(* IEC 61131-3 sources: bevling_machine/framework/sources/02_Devices, 14 files *)

(* ---- F_At.st ---- *)
(* 模块说明：检查设备可用、无忙无故障且位置误差小于 0.01。它检查位置，不检查本次命令序号。 *)
FUNCTION F_At : BOOL
VAR_INPUT
    stStatus : ST_DeviceStatus; (* 本模块对外发布的状态；字段含义见其数据类型。 *)
    lrTarget : LREAL; (* 要检查的目标位置；误差小于 0.01 且设备就绪、无忙无错时返回 TRUE。 *)
END_VAR
FUNCTION F_At : BOOL
(* 位置容差为 0.01 工程单位；这里不做新命令序号校验，用于姿态/互锁判断。 *)
F_At := stStatus.xReady AND NOT stStatus.xBusy
    AND NOT stStatus.xError AND (ABS(stStatus.lrPosition-lrTarget) < 0.01);

(* ---- F_Command.st ---- *)
(* 模块说明：组装设备命令，不执行运动。由设备管理器和对应设备功能块实际处理。 *)
FUNCTION F_Command : ST_DeviceCommand
VAR_INPUT
    eAction : E_DeviceAction; (* 动作类型：无请求、定位、连续运行、点动或停止，见 E_DeviceAction。 *)
    udiID : UDINT; (* 本次命令序号，0 无效；发起新定位时换新序号。 *)
    lrTarget : LREAL; (* 目标工程位置；气缸使用约定的 0/1 端点，连续运行和点动不使用该位置。 *)
    lrVelocity : LREAL; (* 请求速度，单位随设备工程单位定义；尚未完成实机标定。 *)
END_VAR
FUNCTION F_Command : ST_DeviceCommand
(* 只复制字段形成结构体，不等待动作、不直接访问物理设备。 *)
F_Command.eAction := eAction;
F_Command.udiID := udiID;
F_Command.lrTarget := lrTarget;
F_Command.lrVelocity := lrVelocity;

(* ---- F_Done.st ---- *)
(* 模块说明：只有设备完成序号等于本次命令序号、无忙且无故障，才返回动作完成。 *)
FUNCTION F_Done : BOOL
VAR_INPUT
    stStatus : ST_DeviceStatus; (* 本模块对外发布的状态；字段含义见其数据类型。 *)
    udiID : UDINT; (* 本次命令序号，0 无效；发起新定位时换新序号。 *)
END_VAR
FUNCTION F_Done : BOOL
(* 完成必须匹配本次请求；历史 Done 或仅 Busy=FALSE 都不足以作为本步完成条件。 *)
F_Done := (udiID <> 0) AND (stStatus.udiCompletedID = udiID)
    AND NOT stStatus.xBusy AND NOT stStatus.xError;

(* ---- F_NextID.st ---- *)
(* 模块说明：生成本次动作的非零序号。计数到最大值后回到 1，用于排除上一步残留的完成反馈。 *)
FUNCTION F_NextID : UDINT
VAR_IN_OUT
    udiCounter : UDINT; (* 全机共享的动作序号计数器，通过引用传递；由 F_NextID 分配，0 不使用。 *)
END_VAR
FUNCTION F_NextID : UDINT
(* 最大值之后回到 1，跳过无效序号 0；同一机台所有流程共享该计数器。 *)
IF udiCounter = 16#FFFFFFFF THEN udiCounter := 1;
ELSE udiCounter := udiCounter + 1;
END_IF
F_NextID := udiCounter;

(* ---- F_SafetyBypassActive.st ---- *)
(* 模块说明：安全许可软件旁路的唯一判定点。两级开关同时置位才返回 TRUE。 *)
FUNCTION F_SafetyBypassActive : BOOL
VAR_IN_OUT
	stReal : ST_RealDeviceSettings; (* 引用传递，避免每次扫描拷贝整个设置结构体。 *)
END_VAR
FUNCTION F_SafetyBypassActive : BOOL
(* 一级开关与二级确认必须同时置位；任一为 FALSE 就返回 FALSE，保持原有安全逻辑。 *)
F_SafetyBypassActive := stReal.xSafetyBypass AND stReal.xSafetyBypassConfirm;

(* ---- FB_Axis.st ---- *)
(* 模块说明：定位轴适配入口。当前调用内部仿真；真实轴的 MC 功能块、回原点和限位尚未接入。 *)
FUNCTION_BLOCK FB_Axis
VAR_INPUT
    xSimulation : BOOL; (* TRUE 使用内部仿真；当前 FALSE 报未实现 3001，不会接管真实运动。 *)
    xEnable : BOOL; (* 本功能使能，电平有效；失能时不接受新的动作请求。 *)
    xReset : BOOL; (* 故障复位许可；仿真设备仅在故障注入已撤销时清除错误。 *)
    xStall : BOOL; (* 仿真卡住输入；TRUE 暂停位置推进且不发完成，保留忙状态。 *)
    xInjectFault : BOOL; (* 仿真设备故障输入；TRUE 锁存错误码 9001。 *)
    stConfig : ST_DeviceConfig; (* 设备类型、初始位置、软限位与仿真动作时间。 *)
    stCommand : ST_DeviceCommand; (* 当前单设备命令，含动作类型、序号、目标和速度。 *)
END_VAR
VAR_OUTPUT
    stStatus : ST_DeviceStatus; (* 本模块对外发布的状态；字段含义见其数据类型。 *)
END_VAR
VAR
    fbSimulation : FB_SimDevice; (* 内部设备仿真实例，真实设备适配尚未接入。 *)
END_VAR
FUNCTION_BLOCK FB_Axis
(* 真实设备适配尚未接入；关闭仿真时返回 3001，避免误认为已具备实机控制。 *)
fbSimulation(xEnable := xEnable AND xSimulation, xReset := xReset,
    xStall := xStall, xInjectFault := xInjectFault,
    stConfig := stConfig, stCommand := stCommand);
stStatus := fbSimulation.stStatus;
IF NOT xSimulation THEN
    stStatus.xReady := FALSE; stStatus.xBusy := FALSE; stStatus.xActive := FALSE;
    stStatus.xError := TRUE; stStatus.udiErrorID := 3001;
END_IF

(* ---- FB_Cylinder.st ---- *)
(* 模块说明：气缸适配入口。当前用 0/1 位置模拟两端到位；真实电磁阀和到位传感器尚未映射。 *)
FUNCTION_BLOCK FB_Cylinder
VAR_INPUT
    xSimulation : BOOL; (* TRUE 使用内部仿真；当前 FALSE 报未实现 3001，不会接管真实运动。 *)
    xEnable : BOOL; (* 本功能使能，电平有效；失能时不接受新的动作请求。 *)
    xReset : BOOL; (* 故障复位许可；仿真设备仅在故障注入已撤销时清除错误。 *)
    xStall : BOOL; (* 仿真卡住输入；TRUE 暂停位置推进且不发完成，保留忙状态。 *)
    xInjectFault : BOOL; (* 仿真设备故障输入；TRUE 锁存错误码 9001。 *)
    stConfig : ST_DeviceConfig; (* 设备类型、初始位置、软限位与仿真动作时间。 *)
    stCommand : ST_DeviceCommand; (* 当前单设备命令，含动作类型、序号、目标和速度。 *)
END_VAR
VAR_OUTPUT
    stStatus : ST_DeviceStatus; (* 本模块对外发布的状态；字段含义见其数据类型。 *)
END_VAR
VAR
    fbSimulation : FB_SimDevice; (* 内部设备仿真实例，真实设备适配尚未接入。 *)
END_VAR
FUNCTION_BLOCK FB_Cylinder
(* 真实设备适配尚未接入；关闭仿真时返回 3001，避免误认为已具备实机控制。 *)
fbSimulation(xEnable := xEnable AND xSimulation, xReset := xReset,
    xStall := xStall, xInjectFault := xInjectFault,
    stConfig := stConfig, stCommand := stCommand);
stStatus := fbSimulation.stStatus;
IF NOT xSimulation THEN
    stStatus.xReady := FALSE; stStatus.xBusy := FALSE; stStatus.xActive := FALSE;
    stStatus.xError := TRUE; stStatus.udiErrorID := 3001;
END_IF

(* ---- FB_DeviceManager.st ---- *)
FUNCTION_BLOCK FB_DeviceManager
(* 模块说明：统一设备执行入口。首次建立类型和初始位置，每扫描周期按类型调用设备功能块并收集反馈。 *)
VAR_INPUT
	xEnable : BOOL; (* 本功能使能，电平有效；失能时不接受新的动作请求。 *)
	xSimulation : BOOL; (* TRUE 使用内部仿真；当前 FALSE 报未实现 3001，不会接管真实运动。 *)
	xReset : BOOL; (* 故障复位许可；仿真设备仅在故障注入已撤销时清除错误。 *)
	xFaultHold : BOOL; (* 整机故障保持：TRUE 时真实轴强制停车、真实阀失电，直到复位。 *)
	stSim : ST_SimulationSettings; (* 软件仿真设置；设备管理器按设备索引读取卡住与故障注入。 *)
	stReal : ST_RealDeviceSettings; (* 真实设备接管设置；逐台位决定该编号走真实轴还是仿真。 *)
	uiMaterialModel : UINT; (* 当前运行料型 300/450/600；G2 气缸组按此选通其中一个缸下降。 *)
	aCommand : ARRAY[1..17] OF ST_DeviceCommand; (* 统一设备请求数组 1..17；子流程写请求，设备管理器执行。 *)
END_VAR
VAR_OUTPUT
	aStatus : ARRAY[1..17] OF ST_DeviceStatus; (* 各设备的反馈数组 1..17，供判断忙、完成序号、故障和位置。 *)
	aValveOut : ARRAY[1..17] OF BOOL; (* 各设备的阀电气输出电平 1..17；只有已接管的真实气缸可能为 TRUE，供物理映射层取用。 *)
	aValveOutAux : ARRAY[1..17] OF BOOL; (* 第二个执行器的阀电气电平 1..17；当前只有 G1 双压板的 [9] 有效，其余恒 FALSE。 *)
	aG2Valve : ARRAY[1..3] OF BOOL; (* G2 三个侧挡阀的电气电平 1=300，2=450，3=600；未接管时全 FALSE。 *)
	uiG2Band : UINT; (* G2 当前实际下降的料型带号 300/450/600；0 表示三缸全部提升，供诊断观察。 *)
END_VAR
VAR
	aConfig : ARRAY[1..17] OF ST_DeviceConfig; (* 设备配置数组，首扫描按固定编号设置类型和初始姿态。 *)
	aAxis : ARRAY[1..17] OF FB_Axis; (* 定位轴功能块实例数组，只有设备类型为 Axis 的元素被调用。 *)
	aMotor : ARRAY[1..17] OF FB_Motor; (* 连续电机功能块实例数组，供 D1、D3 使用。 *)
	aCylinder : ARRAY[1..17] OF FB_Cylinder; (* 气缸功能块实例数组，按 G 编号驱动对应仿真实例。 *)
	aValve : ARRAY[1..17] OF FB_Valve; (* 阀功能块实例数组，供 G5 喷油及 G6 吹气使用。 *)
	fbRealD1 : FB_RealAxis; (* D1 送料皮带真实轴实例，绑定 songliao。 *)
	fbRealD2 : FB_RealAxis; (* D2 切割走刀真实轴实例，绑定 qiege。 *)
	fbRealD3 : FB_RealAxis; (* D3 盘刀旋转真实轴实例，绑定 pandao（当前按线性模式配置）。 *)
	fbRealD8 : FB_RealAxis; (* D8 平台旋转真实轴实例，绑定 xuanzhuan（台达 ASDA-B3-E）。 *)
	fbRealG1 : FB_RealCylinder; (* G1 下压气缸真实实例，绑定左右两路阀与 G1 两端传感器。 *)
	fbRealG2 : FB_RealCylinderGroup; (* G2 侧挡气缸组真实实例，一台管 300/450/600 三个缸。 *)
	fbRealG3 : FB_RealCylinder; (* G3 侧推气缸真实实例，绑定 xDoG3Valve 与 G3 两端传感器。 *)
	fbRealG9 : FB_RealCylinder; (* G9 盘刀升降真实实例，绑定 xDoG9Valve 与 G9 两端传感器。 *)
	fbRealD6 : FB_RealSensor; (* D6 定长光电真实实例，只读；接管后取代 FB_SimPlant 产生料到位信号。 *)
	axUseReal : ARRAY[1..17] OF BOOL; (* 本扫描逐台接管标志，直接取 stReal.axRealDevice；没有真实实例的编号由回填分支报 3002。 *)
	xBooted : BOOL; (* 本功能块首次初始化完成标志，防止每扫描重写初值。 *)
	i : INT; (* 本扫描数组遍历索引；含义及范围以当前 FOR 循环为准。 *)
END_VAR
FUNCTION_BLOCK FB_DeviceManager
IF NOT xBooted THEN
	(* D1 送料皮带：由真实轴 songliao 承担输送，按定位轴建模（点动/连续运行）。 *)
	aConfig[1].eKind := E_DeviceKind.Axis;
	aConfig[2].eKind := E_DeviceKind.Axis;
	aConfig[3].eKind := E_DeviceKind.Motor;
	aConfig[4].eKind := E_DeviceKind.Axis;
	(* D5 暂按定位升降建模：0=升起避让，1=下降检测，非实际机械坐标。 *)
	aConfig[5].eKind := E_DeviceKind.Axis;
	aConfig[7].eKind := E_DeviceKind.Axis;
	aConfig[8].eKind := E_DeviceKind.Axis;
	FOR i := 9 TO 17 DO aConfig[i].eKind := E_DeviceKind.Cylinder; END_FOR
	aConfig[13].eKind := E_DeviceKind.Valve;
	aConfig[14].eKind := E_DeviceKind.Valve;
	aConfig[12].lrInitialPosition := 1.0;
	FOR i := 1 TO 17 DO
		IF aConfig[i].eKind = E_DeviceKind.Cylinder THEN
			aConfig[i].lrMinPosition := 0.0; aConfig[i].lrMaxPosition := 1.0;
		END_IF
	END_FOR
	(* D2 切割走刀：配方要求 200mm/s、加速度 500；默认 100/50 会把速度削到 100 并拖长加减速段。 *)
	aConfig[2].lrMaxVelocity := 300.0;
	aConfig[2].lrMaxAcceleration := 500.0;
	aConfig[2].lrMaxDeceleration := 500.0;
	xBooted := TRUE;
END_IF

(* 逐台接管标志直接取设置位：是否真的接管由下方回填分支的 CASE 决定。
   新增真实实例时只改 CASE 和实例调用两处，不要再维护第二份白名单。 *)
FOR i := 1 TO 17 DO
	axUseReal[i] := stReal.axRealDevice[i];
END_FOR

(* 四个真实轴实例每扫描必须无条件调用；轴形参写死，无法放进 FOR 循环。
   绑定对照（换电机、改轴名后必须逐行核对：写错不会报编译错误，
   因为任何一个合法轴名都能通过类型检查，只能靠单点测试发现）：
     fbRealD1 -> songliao    设备索引 1，送料皮带（EtherCAT 从站 ASDA_B3_E_CoE_Drive_3）
     fbRealD2 -> qiege       设备索引 2，切割走刀（从站 ASDA_B3_E_CoE_Drive_1）
     fbRealD3 -> pandao      设备索引 3，盘刀旋转（从站 ASDA_B3_E_CoE_Drive_2）
     fbRealD8 -> xuanzhuan   设备索引 8，平台旋转（从站 ASDA_B3_E_CoE_Drive，台达）
   注意：ASDA_B3_E_CoE_Drive_* 是驱动器从站名，代码里写的必须是它下面那个
   轴对象名（songliao/qiege/pandao/xuanzhuan），两者不是一回事。 *)
fbRealD1(Axis := songliao, xUseReal := axUseReal[1], xEnable := xEnable, xReset := xReset,
	xFaultHold := xFaultHold,
	stConfig := aConfig[1], stCommand := aCommand[1], stReal := stReal);
fbRealD2(Axis := qiege, xUseReal := axUseReal[2], xEnable := xEnable, xReset := xReset,
	xFaultHold := xFaultHold,
	stConfig := aConfig[2], stCommand := aCommand[2], stReal := stReal);
fbRealD3(Axis := pandao, xUseReal := axUseReal[3], xEnable := xEnable, xReset := xReset,
	xFaultHold := xFaultHold,
	stConfig := aConfig[3], stCommand := aCommand[3], stReal := stReal);
fbRealD8(Axis := xuanzhuan, xUseReal := axUseReal[8], xEnable := xEnable, xReset := xReset,
	xFaultHold := xFaultHold,
	stConfig := aConfig[8], stCommand := aCommand[8], stReal := stReal);

(* 四个真实气缸实例同样必须无条件调用；传感器与阀逐一对应物理映射符号。
   极性默认 FALSE：传感器高电平有效、阀高电平使能。接线反了只改这里一行，不动流程与互锁。 *)
fbRealG1(xUseReal := axUseReal[9], xEnable := xEnable, xReset := xReset,
	xFaultHold := xFaultHold,
	xSensorRetract := GVL_IO_Physical.xDiG1LRetract, xSensorExtend := GVL_IO_Physical.xDiG1LExtend,
	xSensorRetract2 := GVL_IO_Physical.xDiG1RRetract, xSensorExtend2 := GVL_IO_Physical.xDiG1RExtend,
	xUseSecond := TRUE,
	(* 现场 G1 两只伸出到位传感器已失效：改成只看左右两个缩回信号，两者都无信号并稳定 1s 即认为压到位。
	   传感器修好后把 xExtendByRetract 改回 FALSE 就恢复两端判定，流程和互锁都不用动。 *)
	xExtendByRetract := TRUE, tExtendConfirm := T#1S,
	xInvertSensors := FALSE, xInvertValve := FALSE,
	stConfig := aConfig[9], stCommand := aCommand[9]);
fbRealG2(xUseReal := axUseReal[10], xEnable := xEnable, xReset := xReset,
	xFaultHold := xFaultHold,
	uiMaterialModel := uiMaterialModel,
	xSensorRetract1 := GVL_IO_Physical.xDiG2_300Retract, xSensorExtend1 := GVL_IO_Physical.xDiG2_300Extend,
	xSensorRetract2 := GVL_IO_Physical.xDiG2_450Retract, xSensorExtend2 := GVL_IO_Physical.xDiG2_450Extend,
	xSensorRetract3 := GVL_IO_Physical.xDiG2_600Retract, xSensorExtend3 := GVL_IO_Physical.xDiG2_600Extend,
	xInvertSensors := FALSE, xInvertValve := FALSE,
	stConfig := aConfig[10], stCommand := aCommand[10]);
fbRealG3(xUseReal := axUseReal[11], xEnable := xEnable, xReset := xReset,
	xFaultHold := xFaultHold,
	xSensorRetract := GVL_IO_Physical.xDiG3Retract, xSensorExtend := GVL_IO_Physical.xDiG3Extend,
	xInvertSensors := FALSE, xInvertValve := FALSE,
	stConfig := aConfig[11], stCommand := aCommand[11]);
fbRealG9(xUseReal := axUseReal[17], xEnable := xEnable, xReset := xReset,
	xFaultHold := xFaultHold,
	xSensorRetract := GVL_IO_Physical.xDiG9Retract, xSensorExtend := GVL_IO_Physical.xDiG9Extend,
	xInvertSensors := FALSE, xInvertValve := FALSE,
	stConfig := aConfig[17], stCommand := aCommand[17]);

(* D6 定长光电：只读设备，没有阀也没有动作。
   接线极性反了改 xInvertSensor；光电抖动大改 tDebounce；不需要常亮/常灭监视就把 tStuckTimeout 置 T#0MS。 *)
fbRealD6(xUseReal := axUseReal[6], xEnable := xEnable, xReset := xReset,
	xSensorRaw := GVL_IO_Physical.xDiMaterialLength, xInvertSensor := FALSE,
	tDebounce := T#20MS, tStuckTimeout := T#0MS,
	stConfig := aConfig[6], stCommand := aCommand[6]);

(* 每周期按接管标志二选一：有真实实例的直接回填，否则按设备类型走仿真。
   「实例即事实」：本 CASE 列出全部已实现真实适配的编号，没列到的编号若置了接管位，
   就在 ELSE 分支明确报 3002，避免静默走仿真被误认为已接实机。 *)
(* G2 三个阀默认失电：只有走真实气缸组且缸确实在下降时才会被下面的 CASE 置位。 *)
aG2Valve[1] := FALSE; aG2Valve[2] := FALSE; aG2Valve[3] := FALSE;
uiG2Band := 0;
FOR i := 1 TO 17 DO
	aValveOut[i] := FALSE; aValveOutAux[i] := FALSE;
	IF axUseReal[i] THEN
		CASE i OF
		1: aStatus[i] := fbRealD1.stStatus;
		2: aStatus[i] := fbRealD2.stStatus;
		3: aStatus[i] := fbRealD3.stStatus;
		6: aStatus[i] := fbRealD6.stStatus;
		8: aStatus[i] := fbRealD8.stStatus;
		9: aStatus[i] := fbRealG1.stStatus; aValveOut[i] := fbRealG1.xValve; aValveOutAux[i] := fbRealG1.xValve2;
		10: aStatus[i] := fbRealG2.stStatus; aG2Valve := fbRealG2.aValve; uiG2Band := fbRealG2.uiActiveBand;
		11: aStatus[i] := fbRealG3.stStatus; aValveOut[i] := fbRealG3.xValve;
		17: aStatus[i] := fbRealG9.stStatus; aValveOut[i] := fbRealG9.xValve;
		ELSE
			(* 请求接管但本版本没有对应真实实例：只报错，不启动仿真，保持与老逻辑一致 *)
			aStatus[i].xError := TRUE;
			aStatus[i].udiErrorID := 3002;
		END_CASE
	ELSE
		CASE aConfig[i].eKind OF
		E_DeviceKind.Axis:
			aAxis[i](xSimulation:=xSimulation,xEnable:=xEnable,xReset:=xReset,
				xStall:=stSim.axStall[i],xInjectFault:=stSim.axFault[i],stConfig:=aConfig[i],stCommand:=aCommand[i]);
			aStatus[i] := aAxis[i].stStatus;
		E_DeviceKind.Motor:
			aMotor[i](xSimulation:=xSimulation,xEnable:=xEnable,xReset:=xReset,
				xStall:=stSim.axStall[i],xInjectFault:=stSim.axFault[i],stConfig:=aConfig[i],stCommand:=aCommand[i]);
			aStatus[i] := aMotor[i].stStatus;
		E_DeviceKind.Cylinder:
			aCylinder[i](xSimulation:=xSimulation,xEnable:=xEnable,xReset:=xReset,
				xStall:=stSim.axStall[i],xInjectFault:=stSim.axFault[i],stConfig:=aConfig[i],stCommand:=aCommand[i]);
			aStatus[i] := aCylinder[i].stStatus;
		E_DeviceKind.Valve:
			aValve[i](xSimulation:=xSimulation,xEnable:=xEnable,xReset:=xReset,
				xStall:=stSim.axStall[i],xInjectFault:=stSim.axFault[i],stConfig:=aConfig[i],stCommand:=aCommand[i]);
			aStatus[i] := aValve[i].stStatus;
		END_CASE
	END_IF
END_FOR

(* ---- FB_Motor.st ---- *)
(* 模块说明：连续电机适配入口，供皮带 D1 和盘刀 D3 使用。当前仅仿真运行状态。 *)
FUNCTION_BLOCK FB_Motor
VAR_INPUT
    xSimulation : BOOL; (* TRUE 使用内部仿真；当前 FALSE 报未实现 3001，不会接管真实运动。 *)
    xEnable : BOOL; (* 本功能使能，电平有效；失能时不接受新的动作请求。 *)
    xReset : BOOL; (* 故障复位许可；仿真设备仅在故障注入已撤销时清除错误。 *)
    xStall : BOOL; (* 仿真卡住输入；TRUE 暂停位置推进且不发完成，保留忙状态。 *)
    xInjectFault : BOOL; (* 仿真设备故障输入；TRUE 锁存错误码 9001。 *)
    stConfig : ST_DeviceConfig; (* 设备类型、初始位置、软限位与仿真动作时间。 *)
    stCommand : ST_DeviceCommand; (* 当前单设备命令，含动作类型、序号、目标和速度。 *)
END_VAR
VAR_OUTPUT
    stStatus : ST_DeviceStatus; (* 本模块对外发布的状态；字段含义见其数据类型。 *)
END_VAR
VAR
    fbSimulation : FB_SimDevice; (* 内部设备仿真实例，真实设备适配尚未接入。 *)
END_VAR
FUNCTION_BLOCK FB_Motor
(* 真实设备适配尚未接入；关闭仿真时返回 3001，避免误认为已具备实机控制。 *)
fbSimulation(xEnable := xEnable AND xSimulation, xReset := xReset,
    xStall := xStall, xInjectFault := xInjectFault,
    stConfig := stConfig, stCommand := stCommand);
stStatus := fbSimulation.stStatus;
IF NOT xSimulation THEN
    stStatus.xReady := FALSE; stStatus.xBusy := FALSE; stStatus.xActive := FALSE;
    stStatus.xError := TRUE; stStatus.udiErrorID := 3001;
END_IF

(* ---- FB_RealAxis.st ---- *)
FUNCTION_BLOCK FB_RealAxis
(* 模块说明：真实轴适配层。把统一设备命令翻译成 SoftMotion 动作，并回写与仿真完全一致的接收/完成序号。 *)
VAR_IN_OUT
	Axis : AXIS_REF_SM3; (* 轴节点引用，编译期强制绑定；未接轴无法通过编译，不存在空指针。 *)
END_VAR
VAR_INPUT
	xUseReal : BOOL; (* TRUE 表示本编号由本功能块接管；FALSE 时驱动器保持去使能且不响应任何命令。 *)
	xEnable : BOOL; (* 设备级使能，来自整机许可；FALSE 时主动停止并清序号。 *)
	xReset : BOOL; (* 故障复位，上升沿清锁存错误与 MC 错误。 *)
	stConfig : ST_DeviceConfig; (* 行程、速度、加减速与绝对定位许可。 *)
	stCommand : ST_DeviceCommand; (* 上层统一设备命令，含义与仿真侧完全一致。 *)
	xFaultHold : BOOL; (* 整机故障保持：TRUE 期间强制 MC_Stop 常置并清所有运动请求，直到复位。 *)
	stReal : ST_RealDeviceSettings; (* 相对验证距离、速度与旁路设置。 *)
END_VAR
VAR_OUTPUT
	stStatus : ST_DeviceStatus; (* 与 FB_SimDevice 语义一致，上层无需区分真假设备。 *)
	uiVerifyPhase : UINT; (* 相对验证相位：0 空闲、1 正向、2 停留、3 反向、4 完成、90 中止。 *)
	lrVerifyMeasured : LREAL; (* 本次往返正向段的实测位移，取自轴反馈。 *)
	lrVerifyRatio : LREAL; (* 实测除以指令；只能证明指令与反馈自洽，不能证明单位就是毫米。 *)
END_VAR
VAR
	fbPower : MC_Power; (* 伺服使能，接管期间保持上电。 *)
	fbReset : MC_Reset; (* 清 MC 错误。 *)
	fbStop : MC_Stop; (* 受控停止，停止请求需保持到 Done。 *)
	fbMoveAbs : MC_MoveAbsolute; (* 绝对定位，仅在 xAbsoluteAllowed 为 TRUE 时使用。 *)
	fbMoveRel : MC_MoveRelative; (* 相对定位，验证模式的两段行程使用。 *)
	fbMoveVel : MC_MoveVelocity; (* 连续运行与点动共用，两者相位互斥；方向必须显式给出。 *)
	fbHoming : CmpHCMotion.MC_Homing; (* 上位机回零：由 PLC 自己按轴配置的回零方式走，不依赖驱动器支持 DS402 回零。 *)
	fbReadPos : MC_ReadActualPosition; (* 实际位置反馈。 *)
	fbReadStatus : MC_ReadStatus; (* 轴状态，用于判断故障停止。 *)
	fbReadErr : MC_ReadAxisError; (* 轴错误码，供在线排查。 *)
	rtReset : R_TRIG; (* 复位上升沿。 *)
	tonEnable : TON; (* 命令已接收但轴未使能的 3 秒超时。 *)
	tonDwell : TON; (* 验证往返之间的停留，保证 Execute 拉低形成新上升沿。 *)
	tonHome : TON; (* 回零超时；找不到原点时按 2004 暴露，避免无限等待。 *)
	udiLastID : UDINT; (* 上次已接受序号，用于识别新命令。 *)
	udiActiveID : UDINT; (* 正在执行的序号，完成时回写。 *)
	xPending : BOOL; (* 已接收但尚未启动，等待轴使能。 *)
	xStopLatch : BOOL; (* 停止请求锁存，保持到 MC_Stop 完成。 *)
	xStopReq : BOOL; (* 本扫描停止请求。 *)
	xMoveAbsReq : BOOL; (* 本扫描绝对定位请求。 *)
	xMoveRelReq : BOOL; (* 本扫描相对定位请求。 *)
	xMoveVelReq : BOOL; (* 本扫描速度模式请求，连续运行与点动共用。 *)
	xHomeReq : BOOL; (* 本扫描回零请求，保持到 Done。 *)
	xHomed : BOOL; (* 本次上电后已成功回零；成功后允许绝对定位，断电或重新下载后清零。 *)
	uiPhase : UINT; (* 动作相位：0 空闲、10 等待使能、20 绝对、30/31/32 验证三段、40 连续、50 点动、60 回零、90 中止。 *)
	lrVerifyStart : LREAL; (* 验证正向段起点位置。 *)
	lrRelDistance : LREAL; (* 本次相对定位距离，正负决定方向。 *)
	lrRelVelocity : LREAL; (* 本次相对定位速度，取正值。 *)
	lrCmdVelocity : LREAL; (* 连续运行与点动的限幅后速度，带符号。 *)
END_VAR
FUNCTION_BLOCK FB_RealAxis
(* ===== 1. 读取块无条件调用，保证反馈新鲜 ===== *)
fbReadPos(Axis := Axis, Enable := TRUE);
fbReadStatus(Axis := Axis, Enable := TRUE);
fbReadErr(Axis := Axis, Enable := TRUE);
rtReset(CLK := xReset);

stStatus.lrPosition := fbReadPos.Position;
stStatus.xRealActive := xUseReal;

(* ===== 2. 复位：只在接管状态下响应，避免误清其它轴 ===== *)
IF xUseReal AND rtReset.Q THEN
	stStatus.xError := FALSE;
	stStatus.udiErrorID := 0;
	xStopLatch := FALSE;
	xPending := FALSE;
	uiPhase := 0;
	uiVerifyPhase := 0;
	udiLastID := 0;
	udiActiveID := 0;
	stStatus.udiAcceptedID := 0;
	stStatus.udiCompletedID := 0;
	stStatus.xBusy := FALSE;
	stStatus.xActive := FALSE;
END_IF

(* ===== 3. 定时器：用上扫描状态驱动，避免与状态判定循环依赖 ===== *)
tonEnable(IN := xPending AND xUseReal, PT := T#3S);
tonDwell(IN := (uiPhase = 31), PT := stReal.tVerifyDwell);
tonHome(IN := (uiPhase = 60), PT := stReal.tHomeTimeout);

(* ===== 4. 请求默认全部撤销 ===== *)
xStopReq := FALSE;
xMoveAbsReq := FALSE;
xMoveRelReq := FALSE;
xMoveVelReq := FALSE;
xHomeReq := FALSE;
lrRelDistance := 0.0;
lrRelVelocity := 0.0;
lrCmdVelocity := 0.0;

(* ===== 4.5 整机故障保持：故障期间主动停车，不依赖 xPermit 间接撤销 ===== *)
(* 为什么需要：进入 Fault 时上层只是让 xPermit 变 FALSE，请求被换成 Stop。但 Stop 是
   一次性的动作请求，盘刀这类连续运行设备在 MC_Stop 完成后再无后续指令，表现就是
   “PLC 认为已停、实际还在转”。这里改用 xFaultHold 强制 MC_Stop 常置，直到真正复位。 *)
IF xFaultHold THEN
	xStopReq := TRUE;
	xPending := FALSE;
	xMoveAbsReq := FALSE; xMoveRelReq := FALSE; xMoveVelReq := FALSE; xHomeReq := FALSE;
	uiPhase := 0; uiVerifyPhase := 0;
	udiLastID := 0; udiActiveID := 0;
	stStatus.udiAcceptedID := 0; stStatus.udiCompletedID := 0;
	stStatus.xBusy := FALSE; stStatus.xActive := FALSE;
END_IF

(* ===== 5. 主状态判定 ===== *)
IF NOT xUseReal THEN
	(* 未接管：不产生任何运动请求，驱动器由 MC_Power 去使能。 *)
	xPending := FALSE; xStopLatch := FALSE;
	uiPhase := 0; uiVerifyPhase := 0;
	udiLastID := 0; udiActiveID := 0;
	stStatus.xReady := FALSE;
	stStatus.xBusy := FALSE; stStatus.xActive := FALSE;
	stStatus.udiAcceptedID := 0; stStatus.udiCompletedID := 0;
	stStatus.xError := FALSE; stStatus.udiErrorID := 0;
ELSIF xFaultHold THEN
	(* 故障保持：只允许停止，不接收新命令，也不发布就绪。 *)
	stStatus.xReady := FALSE;
	stStatus.xBusy := FALSE; stStatus.xActive := FALSE;
	stStatus.udiAcceptedID := 0; stStatus.udiCompletedID := 0;
ELSE
	(* --- 5.1 接收新序号：新序号就是新命令，不用边沿检测 --- *)
	IF (stCommand.udiID <> 0) AND (stCommand.udiID <> udiLastID)
		AND xEnable AND NOT stStatus.xError THEN
		udiLastID := stCommand.udiID;
		udiActiveID := udiLastID;
		stStatus.udiAcceptedID := udiActiveID;
		stStatus.udiCompletedID := 0;
		stStatus.xBusy := TRUE; stStatus.xActive := FALSE;
		uiVerifyPhase := 0;
		xPending := TRUE;
		uiPhase := 10;
		xStopLatch := FALSE;
	END_IF

	(* --- 5.2 停止请求锁存：保持到 MC_Stop 完成，不能提前撤 Execute --- *)
	IF (stCommand.eAction = E_DeviceAction.Stop) OR (NOT xEnable) THEN
		(* 只在真的有动作时才锁存，避免 Stop 常驻时每扫描重复触发 MC_Stop。 *)
		IF xPending OR (uiPhase <> 0) THEN xStopLatch := TRUE; END_IF
	ELSIF (stCommand.eAction = E_DeviceAction.None) AND (uiPhase <> 0) THEN
		xStopLatch := TRUE;
	END_IF
	IF fbStop.Done THEN xStopLatch := FALSE; END_IF

	IF xStopLatch THEN
		xStopReq := TRUE;
		xPending := FALSE;
		uiPhase := 0; uiVerifyPhase := 0;
		udiLastID := 0; udiActiveID := 0;
		stStatus.udiAcceptedID := 0; stStatus.udiCompletedID := 0;
		stStatus.xBusy := FALSE; stStatus.xActive := FALSE;
	ELSIF xPending THEN
		(* --- 5.3 等轴使能；就绪后按动作类型进入相位，3 秒未使能报 2003 --- *)
		IF fbPower.Status THEN
			xPending := FALSE;
			CASE stCommand.eAction OF
			E_DeviceAction.Position:
				(* 已回零优先走绝对定位：相对验证只是未回零时的临时替代，回零成功后不再需要。 *)
				IF xHomed OR stConfig.xAbsoluteAllowed THEN
					uiPhase := 20;
				ELSIF stReal.xRelativeVerify THEN
					lrVerifyStart := fbReadPos.Position;
					uiPhase := 30; uiVerifyPhase := 1;
				ELSE
					(* 未回零不允许绝对定位：报 2002 且不置完成位，由上层按步号超时暴露。 *)
					stStatus.xError := TRUE; stStatus.udiErrorID := 2002;
					uiPhase := 0; uiVerifyPhase := 0;
				END_IF
			E_DeviceAction.Run:
				uiPhase := 40;
			E_DeviceAction.Jog:
				uiPhase := 50;
			E_DeviceAction.Home:
				uiPhase := 60;
			ELSE
				uiPhase := 0;
			END_CASE
		ELSIF tonEnable.Q THEN
			xPending := FALSE; uiPhase := 0;
			stStatus.xError := TRUE; stStatus.udiErrorID := 2003;
			stStatus.xBusy := FALSE;
		END_IF
	END_IF

	(* --- 5.4 按相位生成限幅后的运动参数 --- *)
	CASE uiPhase OF
	30:
		lrRelDistance := LIMIT(0.0, stReal.lrVerifyDistance, 20.0);
		lrRelVelocity := LIMIT(0.01, stReal.lrVerifyVelocity, stConfig.lrMaxVelocity);
	32:
		lrRelDistance := -LIMIT(0.0, stReal.lrVerifyDistance, 20.0);
		lrRelVelocity := LIMIT(0.01, stReal.lrVerifyVelocity, stConfig.lrMaxVelocity);
	40:
		(* 连续运行：按设备配置限幅，不使用验证低速。 *)
		lrCmdVelocity := LIMIT(-stConfig.lrMaxVelocity, stCommand.lrVelocity, stConfig.lrMaxVelocity);
	50:
		(* 点动：用设备最大速度与手动上限 lrManualVelocityMax 的较小者限幅；不能再用验证速度，否则手动最高只有 2mm/s。 *)
		lrCmdVelocity := LIMIT(0.01, ABS(stCommand.lrVelocity),
			MIN(stConfig.lrMaxVelocity, stReal.lrManualVelocityMax));
		IF stCommand.lrVelocity < 0.0 THEN lrCmdVelocity := -lrCmdVelocity; END_IF
	END_CASE

	xMoveAbsReq := (uiPhase = 20);
	xMoveRelReq := (uiPhase = 30) OR (uiPhase = 32);
	xMoveVelReq := (uiPhase = 40) OR (uiPhase = 50);
	xHomeReq := (uiPhase = 60);
END_IF

(* ===== 6. MC 块无条件调用：漏调用会报 SMC_FB_WASNT_CALLED_DURING_MOTION ===== *)
fbPower(Axis := Axis, Enable := xUseReal AND xEnable,
	bRegulatorOn := xUseReal AND xEnable, bDriveStart := xUseReal AND xEnable);
fbReset(Axis := Axis, Execute := xUseReal AND rtReset.Q);
fbStop(Axis := Axis, Execute := xStopReq OR xFaultHold, Deceleration := stConfig.lrMaxDeceleration);
fbMoveRel(Axis := Axis, Execute := xMoveRelReq, Distance := lrRelDistance,
	Velocity := lrRelVelocity, Acceleration := stConfig.lrMaxAcceleration,
	Deceleration := stConfig.lrMaxDeceleration);
fbMoveAbs(Axis := Axis, Execute := xMoveAbsReq, Position := stCommand.lrTarget,
	Velocity := LIMIT(0.01, ABS(stCommand.lrVelocity), stConfig.lrMaxVelocity),
	Acceleration := stConfig.lrMaxAcceleration, Deceleration := stConfig.lrMaxDeceleration);
fbMoveVel(Axis := Axis, Execute := xMoveVelReq,
	Velocity := ABS(lrCmdVelocity),
	Direction := SEL(lrCmdVelocity < 0.0, MC_Direction.positive, MC_Direction.negative),
	Acceleration := stConfig.lrMaxAcceleration,
	Deceleration := stConfig.lrMaxDeceleration);
(* 回零走 MC_Homing（上位机回零）：回零方式、开始方向、零点信号、快慢速全部来自轴配置，
   本块只给 Axis 和 Execute。驱动器不支持 DS402 回零，用 MC_Home 会一直卡在 Homing 状态不动。 *)
fbHoming(Axis := Axis, Execute := xHomeReq);

(* ===== 7. 完成判定与序号回写 ===== *)
IF xUseReal THEN
	CASE uiPhase OF
	20:
		IF fbMoveAbs.Done THEN
			stStatus.udiCompletedID := udiActiveID;
			stStatus.xBusy := FALSE; stStatus.xActive := FALSE;
			uiPhase := 0;
		ELSIF fbMoveAbs.CommandAborted THEN
			stStatus.xBusy := FALSE; uiPhase := 0;
		END_IF
	30:
		IF fbMoveRel.Done THEN
			lrVerifyMeasured := fbReadPos.Position - lrVerifyStart;
			uiPhase := 31; uiVerifyPhase := 2;
		ELSIF fbMoveRel.CommandAborted THEN
			uiPhase := 90; uiVerifyPhase := 90;
			stStatus.xError := TRUE; stStatus.udiErrorID := 2005;
			stStatus.xBusy := FALSE;
		END_IF
	31:
		IF tonDwell.Q THEN
			uiPhase := 32; uiVerifyPhase := 3;
		END_IF
	32:
		IF fbMoveRel.Done THEN
			IF stReal.lrVerifyDistance > 0.001 THEN
				lrVerifyRatio := lrVerifyMeasured / stReal.lrVerifyDistance;
			END_IF
			uiPhase := 0; uiVerifyPhase := 4;
			stStatus.udiCompletedID := udiActiveID;
			stStatus.xBusy := FALSE; stStatus.xActive := FALSE;
		ELSIF fbMoveRel.CommandAborted THEN
			uiPhase := 90; uiVerifyPhase := 90;
			stStatus.xError := TRUE; stStatus.udiErrorID := 2005;
			stStatus.xBusy := FALSE;
		END_IF
	40:
		(* 连续运行：建立速度后回写完成位，但保持相位直到命令改变。 *)
		IF fbMoveVel.InVelocity THEN
			stStatus.xActive := TRUE;
			stStatus.xBusy := FALSE;
			stStatus.udiCompletedID := udiActiveID;
		END_IF
	50:
		(* 点动：与仿真一致，不置完成位，靠松开后的 None/Stop 停止。 *)
		stStatus.xActive := fbMoveVel.InVelocity;
		stStatus.xBusy := TRUE;
	60:
		(* 回零：Done 后置 xHomed 并放行绝对定位；超时报 2004 且不置完成位，避免上层误判已到位。 *)
		IF fbHoming.Done THEN
			xHomed := TRUE;
			stStatus.udiCompletedID := udiActiveID;
			stStatus.xBusy := FALSE; stStatus.xActive := FALSE;
			uiPhase := 0;
		ELSIF fbHoming.CommandAborted THEN
			(* 被其它运动块打断：只清忙标志退出相位，既不置完成位也不置故障，由上层按步号超时暴露。 *)
			stStatus.xBusy := FALSE; uiPhase := 0;
		ELSIF tonHome.Q THEN
			xHomed := FALSE;
			stStatus.xError := TRUE; stStatus.udiErrorID := 2004;
			stStatus.xBusy := FALSE; uiPhase := 0;
		END_IF
	END_CASE

	(* --- MC 错误汇总：只锁存第一条，40000 为前缀，低 16 位保留原码便于查手册 --- *)
	IF NOT stStatus.xError THEN
		IF fbPower.Error THEN
			stStatus.xError := TRUE; stStatus.udiErrorID := UDINT#40000 + TO_UDINT(fbPower.ErrorID);
		ELSIF fbReset.Error THEN
			stStatus.xError := TRUE; stStatus.udiErrorID := UDINT#40000 + TO_UDINT(fbReset.ErrorID);
		ELSIF fbStop.Error THEN
			stStatus.xError := TRUE; stStatus.udiErrorID := UDINT#40000 + TO_UDINT(fbStop.ErrorID);
		ELSIF fbMoveRel.Error THEN
			stStatus.xError := TRUE; stStatus.udiErrorID := UDINT#40000 + TO_UDINT(fbMoveRel.ErrorID);
		ELSIF fbMoveAbs.Error THEN
			stStatus.xError := TRUE; stStatus.udiErrorID := UDINT#40000 + TO_UDINT(fbMoveAbs.ErrorID);
		ELSIF fbMoveVel.Error THEN
			stStatus.xError := TRUE; stStatus.udiErrorID := UDINT#40000 + TO_UDINT(fbMoveVel.ErrorID);
		ELSIF fbHoming.Error THEN
			stStatus.xError := TRUE; stStatus.udiErrorID := UDINT#40000 + TO_UDINT(fbHoming.ErrorID);
		END_IF
	END_IF
END_IF

(* ===== 8. 就绪与故障收尾 ===== *)
stStatus.xReady := xUseReal AND xEnable AND NOT stStatus.xError;
stStatus.xHomed := xUseReal AND xHomed;
IF stStatus.xError THEN
	stStatus.xBusy := FALSE;
	stStatus.xActive := FALSE;
END_IF

(* ---- FB_RealCylinder.st ---- *)
FUNCTION_BLOCK FB_RealCylinder
(* 模块说明：真实气缸适配层。读取两端到位传感器判定姿态，按统一设备命令驱动单电控阀，
   回写与 FB_SimDevice 完全一致的接收/完成序号，使上层流程与互锁无需区分真假气缸。
   某个端点传感器损坏时用 xExtendByRetract 退让：只看缩回信号，全部消失并稳定后视为伸出到位。 *)
VAR_INPUT
	xUseReal : BOOL; (* TRUE 表示本编号由真实气缸接管；FALSE 时阀保持失电且不响应任何命令。 *)
	xEnable : BOOL; (* 设备级使能，来自整机许可；FALSE 时阀失电并清序号。 *)
	xReset : BOOL; (* 故障复位上升沿；清锁存错误并允许重新建立姿态。 *)
	xSensorRetract : BOOL; (* 缩回到位传感器原始电平，TRUE 表示该端有信号。 *)
	xSensorExtend : BOOL; (* 伸出到位传感器原始电平，TRUE 表示该端有信号。 *)
	xSensorRetract2 : BOOL; (* 第二组（右压板）缩回到位原始电平；仅 xUseSecond 为 TRUE 时参与判定。 *)
	xSensorExtend2 : BOOL; (* 第二组（右压板）伸出到位原始电平；仅 xUseSecond 为 TRUE 时参与判定。 *)
	xUseSecond : BOOL := FALSE; (* TRUE 表示由两个同步执行器组成：两组传感器必须同时到位才算该端到位。 *)
	xExtendByRetract : BOOL := FALSE; (* 退让模式：伸出端传感器不可用时置 TRUE，改用「所有缩回信号都消失」推断伸出到位；默认 FALSE 仍按两端判定。 *)
	tExtendConfirm : TIME := T#1S; (* 仅退让模式有效：缩回信号消失并持续该时间才确认伸出到位，避免气缸刚起步就误判为已伸出。 *)
	xInvertSensors : BOOL; (* TRUE 表示两个传感器接线为低电平有效，本层统一取反，不动上层。 *)
	xInvertValve : BOOL; (* TRUE 表示阀为低电平使能；默认 FALSE，即高电平使能。 *)
	xFaultHold : BOOL := FALSE; (* 整机故障保持：TRUE 时阀立即失电并撤销保位，直到复位。 *)
	tSensorTimeout : TIME := T#3S; (* 两端均无信号达到该时间判为传感器丢失，报 3004；双执行器时也包含两侧不同步。 *)
	tTravelTimeout : TIME := T#10S; (* 命令发出后未到位达到该时间判为动作超时，报 3005。 *)
	stConfig : ST_DeviceConfig; (* 行程范围，语义与仿真侧一致；气缸只使用 0/1 两端。 *)
	stCommand : ST_DeviceCommand; (* 上层统一设备命令，气缸只响应 Position 的 0/1 目标。 *)
END_VAR
VAR_OUTPUT
	stStatus : ST_DeviceStatus; (* 与 FB_SimDevice 语义一致；lrPosition 取 0.0 缩回、1.0 伸出。 *)
	xValve : BOOL; (* 阀电气输出电平，已含 xInvertValve；直接接物理输出点。 *)
	xValve2 : BOOL; (* 第二个执行器的阀电气输出电平；xUseSecond 为 FALSE 时恒为 FALSE。 *)
END_VAR
VAR
	rtReset : R_TRIG; (* 复位上升沿。 *)
	tonNoSensor : TON; (* 两端均无信号的持续计时。 *)
	tonExtendConfirm : TON; (* 退让模式下「缩回信号全部消失」的持续计时，到时才确认伸出到位。 *)
	tonTravel : TON; (* 命令发出后等待到位的计时。 *)
	udiLastID : UDINT; (* 上次已接受的命令序号。 *)
	xSenseRetract : BOOL; (* 取反处理后的缩回信号：双执行器时为两侧 AND，TRUE 表示两侧都缩回到位。 *)
	xRetractAny : BOOL; (* 取反处理后的缩回信号：双执行器时为两侧 OR，TRUE 表示至少一侧仍停在缩回位。退让模式用它判「两侧都离开」。 *)
	xSenseExtend : BOOL; (* 取反处理后的伸出信号。 *)
	xPositionKnown : BOOL; (* 姿态是否已由传感器确立；未确立时 xReady 必须为 FALSE，防止上层把未知当成已缩回。 *)
	lrLastKnown : LREAL; (* 最后一次确立的姿态；传感器全灭时保持该值。 *)
	xCmdValid : BOOL; (* 当前存在有效的保位命令，阀按此持续输出。 *)
	xCmdExtend : BOOL; (* 有效命令期望的端点：TRUE 伸出，FALSE 缩回。 *)
	xTravelling : BOOL; (* 尚未确认到达目标端点。 *)
END_VAR
FUNCTION_BLOCK FB_RealCylinder
rtReset(CLK := xReset);

(* ===== 1. 复位：只清错误与序号，姿态仍由传感器决定 ===== *)
IF xUseReal AND rtReset.Q THEN
	stStatus.xError := FALSE; stStatus.udiErrorID := 0;
	xCmdValid := FALSE; xTravelling := FALSE; udiLastID := 0;
	stStatus.udiAcceptedID := 0; stStatus.udiCompletedID := 0;
	tonNoSensor(IN := FALSE);
	tonTravel(IN := FALSE);
END_IF

(* ===== 2. 传感器取反与姿态判定 ===== *)
xSenseRetract := xSensorRetract XOR xInvertSensors;
xSenseExtend := xSensorExtend XOR xInvertSensors;

(* 双执行器：两组必须同时到位才算该端到位。
   左侧在上、右侧在下时两个都为 FALSE，自然落进下面的“两端都无信号”分支：
   保持上次姿态，持续 tSensorTimeout 才报 3004，与单缸中间态同一套处理。
   同时另算一个 OR 合成量给退让模式用：AND 取反只能得到「至少一侧离开」，
   而退让模式要的是「两侧都离开」，所以必须在合并之前留一份单侧信号。 *)
xRetractAny := xSenseRetract;
IF xUseSecond THEN
	xRetractAny := xRetractAny OR (xSensorRetract2 XOR xInvertSensors);
	xSenseRetract := xSenseRetract AND (xSensorRetract2 XOR xInvertSensors);
	xSenseExtend := xSenseExtend AND (xSensorExtend2 XOR xInvertSensors);
END_IF

(* 退让模式：伸出端传感器不可用，只认缩回信号。
   判定 = 左右两侧都没有缩回信号（都离开缩回位）并持续 tExtendConfirm；
   必须延时确认：缩回信号在气缸刚起步就掉，不延时会在压板还没压下去时就报已伸出，
   上层的压紧判定和自动流程会提前放行。延时期间保持上次姿态。 *)
tonExtendConfirm(IN := xUseReal AND xExtendByRetract AND NOT xRetractAny, PT := tExtendConfirm);
IF xExtendByRetract THEN
	xSenseExtend := tonExtendConfirm.Q;
END_IF

(* 退让模式下「两端都无信号」正是伸出到位的正常表现，不能再按传感器丢失报 3004，所以此模式关闭该计时。 *)
tonNoSensor(IN := xUseReal AND NOT xExtendByRetract AND NOT xSenseRetract AND NOT xSenseExtend, PT := tSensorTimeout);

IF xSenseRetract AND xSenseExtend THEN
	(* 两端同时有信号：传感器短路、磁环位置错或机械卡在中间，姿态不可信 *)
	xPositionKnown := FALSE;
	stStatus.lrPosition := lrLastKnown;
	stStatus.xError := TRUE; stStatus.udiErrorID := 3003;
ELSIF xSenseExtend THEN
	xPositionKnown := TRUE; lrLastKnown := 1.0; stStatus.lrPosition := 1.0;
ELSIF xSenseRetract THEN
	xPositionKnown := TRUE; lrLastKnown := 0.0; stStatus.lrPosition := 0.0;
ELSE
	(* 两端都没有信号：保持最后姿态；从未确立过则 xReady 一直为 FALSE *)
	stStatus.lrPosition := lrLastKnown;
	IF tonNoSensor.Q AND NOT stStatus.xError THEN
		xPositionKnown := FALSE;
		stStatus.xError := TRUE; stStatus.udiErrorID := 3004;
	END_IF
END_IF

(* ===== 3. 命令接收与保位判定 ===== *)
IF NOT xUseReal THEN
	(* 未接管：不驱动阀，也不发布就绪，避免被上层当成可用设备 *)
	xCmdValid := FALSE; xTravelling := FALSE; udiLastID := 0;
	stStatus.xReady := FALSE; stStatus.xBusy := FALSE; stStatus.xActive := FALSE;
	stStatus.udiAcceptedID := 0; stStatus.udiCompletedID := 0;
ELSIF NOT xEnable OR stStatus.xError OR xFaultHold THEN
	(* 故障或整机故障保持时阀失电，不带错误继续动作 *)
	xCmdValid := FALSE; xTravelling := FALSE;
	stStatus.xReady := FALSE; stStatus.xBusy := FALSE; stStatus.xActive := FALSE;
ELSE
	stStatus.xReady := xEnable AND xPositionKnown;

	(* 新序号即新命令；姿态未确立时不接受，防止朝未知状态动作 *)
	IF (stCommand.udiID <> 0) AND (stCommand.udiID <> udiLastID)
		AND xEnable AND xPositionKnown AND NOT stStatus.xBusy THEN
		udiLastID := stCommand.udiID;
		stStatus.udiAcceptedID := udiLastID; stStatus.udiCompletedID := 0;
		CASE stCommand.eAction OF
		E_DeviceAction.Position:
			IF (stCommand.lrTarget < stConfig.lrMinPosition - 0.01)
				OR (stCommand.lrTarget > stConfig.lrMaxPosition + 0.01) THEN
				stStatus.xError := TRUE; stStatus.udiErrorID := 2001;
				xCmdValid := FALSE;
			ELSE
				xCmdExtend := stCommand.lrTarget > 0.5;
				xCmdValid := TRUE;
				xTravelling := TRUE;
				stStatus.xBusy := TRUE;
			END_IF
		E_DeviceAction.Stop, E_DeviceAction.None:
			xCmdValid := FALSE; xTravelling := FALSE;
			stStatus.udiAcceptedID := 0; stStatus.udiCompletedID := 0;
			udiLastID := 0;
		ELSE
			(* 气缸没有连续运行、点动和回零，明确报错而不是静默不动 *)
			stStatus.xError := TRUE; stStatus.udiErrorID := 2001;
			xCmdValid := FALSE;
		END_CASE
	END_IF

	(* 命令被撤销或失能：立即取消保位，阀随之失电 *)
	IF (stCommand.eAction = E_DeviceAction.Stop) OR (stCommand.eAction = E_DeviceAction.None)
		OR NOT xEnable THEN
		xCmdValid := FALSE; xTravelling := FALSE;
		stStatus.xBusy := FALSE;
	END_IF

	(* 到位判定：姿态已知且与命令期望的端点一致即算完成 *)
	IF xCmdValid AND xPositionKnown THEN
		IF (xCmdExtend AND (stStatus.lrPosition > 0.5))
			OR ((NOT xCmdExtend) AND (stStatus.lrPosition < 0.5)) THEN
			IF xTravelling THEN stStatus.udiCompletedID := udiLastID; END_IF
			xTravelling := FALSE;
			stStatus.xBusy := FALSE;
		END_IF
	END_IF
END_IF

(* ===== 4. 到位超时 ===== *)
tonTravel(IN := xUseReal AND xTravelling AND xCmdValid, PT := tTravelTimeout);
IF tonTravel.Q AND NOT stStatus.xError THEN
	stStatus.xError := TRUE; stStatus.udiErrorID := 3005;
	stStatus.xBusy := FALSE;
	xTravelling := FALSE;
END_IF

(* ===== 5. 阀输出：按保位命令持续输出，不是只在动作过程中输出 ===== *)
xValve := FALSE;
xValve2 := FALSE;
IF xCmdValid AND xUseReal AND NOT stStatus.xError AND NOT xFaultHold THEN
	xValve := xCmdExtend;
	IF xUseSecond THEN xValve2 := xCmdExtend; END_IF
END_IF
IF xInvertValve THEN xValve := NOT xValve; END_IF
IF xInvertValve AND xUseSecond THEN xValve2 := NOT xValve2; END_IF

(* ===== 6. 收尾 ===== *)
stStatus.xReady := stStatus.xReady AND xUseReal AND NOT stStatus.xError;
stStatus.xActive := xCmdValid;
(* 气缸没有回零动作，用“姿态已确立”代替，供整机统计已接管设备是否可信 *)
stStatus.xHomed := xUseReal AND xPositionKnown;

(* ---- FB_RealCylinderGroup.st ---- *)
FUNCTION_BLOCK FB_RealCylinderGroup
(* 模块说明：按料型选通的真实气缸组适配层（G2 侧挡用，300/450/600 三缸共用设备索引 10）。
   同一时刻只允许一个气缸下降，其余两个强制提升；回写与 FB_SimDevice 完全一致的接收/完成序号，
   使上层流程与互锁无需区分单缸、多缸或仿真。
   命令目标 lrTarget：0 = 三缸全部提升；300 / 450 / 600 = 对应料型气缸下降，其余两个提升。
   lrTarget 在 0..1 之间时按单缸旧语义映射：>0.5 视为「降到当前料型」，<=0.5 视为三缸全部提升。 *)
VAR_INPUT
	xUseReal : BOOL; (* TRUE 表示本编号由真实气缸组接管；FALSE 时三个阀全部失电且不响应任何命令。 *)
	xEnable : BOOL; (* 设备级使能，来自整机许可；FALSE 时阀失电并清序号。 *)
	xReset : BOOL; (* 故障复位上升沿；清锁存错误与序号。 *)
	xFaultHold : BOOL; (* 整机故障保持：TRUE 时三个阀立即失电，直到复位。 *)
	uiMaterialModel : UINT; (* 当前运行料型 300/450/600；旧语义 lrTarget>0.5 时降到本料型。 *)
	xSensorRetract1 : BOOL; (* 1 号缸（300）提升到位传感器原始电平，TRUE 表示该端有信号。 *)
	xSensorExtend1 : BOOL; (* 1 号缸（300）下降到位传感器原始电平。 *)
	xSensorRetract2 : BOOL; (* 2 号缸（450）提升到位传感器原始电平。 *)
	xSensorExtend2 : BOOL; (* 2 号缸（450）下降到位传感器原始电平。 *)
	xSensorRetract3 : BOOL; (* 3 号缸（600）提升到位传感器原始电平。 *)
	xSensorExtend3 : BOOL; (* 3 号缸（600）下降到位传感器原始电平。 *)
	xInvertSensors : BOOL; (* TRUE 表示六个传感器均为低电平有效，本层统一取反，不动上层。 *)
	xInvertValve : BOOL; (* TRUE 表示三个阀均为低电平使能；默认 FALSE，即高电平使能。 *)
	tSensorTimeout : TIME := T#3S; (* 六个传感器全部无信号达到该时间判为整组丢失，报 3004。 *)
	tTravelTimeout : TIME := T#10S; (* 命令发出后目标姿态未达成达到该时间判为动作超时，报 3005。 *)
	stConfig : ST_DeviceConfig; (* 行程范围，语义与仿真侧一致；组内气缸只使用 0/1 两端。 *)
	stCommand : ST_DeviceCommand; (* 上层统一设备命令，本层只响应 Position 的 0/300/450/600 目标。 *)
END_VAR
VAR_OUTPUT
	stStatus : ST_DeviceStatus; (* 与 FB_SimDevice 语义一致；目标缸下降到位 1.0，三缸全提 0.0，中间保持上次值。 *)
	aValve : ARRAY[1..3] OF BOOL; (* 三个阀的电气电平（已含 xInvertValve），直接接物理输出点；索引 1=300，2=450，3=600。 *)
	uiActiveBand : UINT; (* 当前实际下降的料型带号；0 表示三个缸都在提升位。 *)
END_VAR
VAR
	rtReset : R_TRIG; (* 复位上升沿。 *)
	tonNoSensor : TON; (* 六个传感器全部无信号的持续计时。 *)
	tonTravel : TON; (* 命令发出后等待到位的计时。 *)
	udiLastID : UDINT; (* 上次已接受的命令序号。 *)
	aRetract : ARRAY[1..3] OF BOOL; (* 取反处理后的三路提升信号。 *)
	aExtend : ARRAY[1..3] OF BOOL; (* 取反处理后的三路下降信号。 *)
	xAllRetract : BOOL; (* 三个缸都确认在提升位。 *)
	xPositionKnown : BOOL; (* 三缸姿态是否都已由传感器确立；未确立时 xReady 必须为 FALSE，防止上层把未知当成已提升。 *)
	xCmdValid : BOOL; (* 当前存在有效的保位命令，阀按此持续输出。 *)
	uiTargetBand : UINT; (* 有效命令期望下降的料型带号；0 表示三缸全部提升。 *)
	xTravelling : BOOL; (* 尚未确认到达命令要求的姿态。 *)
	i : INT; (* 本扫描数组遍历索引；含义及范围以当前 FOR 循环为准。 *)
END_VAR
FUNCTION_BLOCK FB_RealCylinderGroup
rtReset(CLK := xReset);

(* ===== 1. 复位：只清错误与序号，姿态仍由传感器决定 ===== *)
IF xUseReal AND rtReset.Q THEN
	stStatus.xError := FALSE; stStatus.udiErrorID := 0;
	xCmdValid := FALSE; xTravelling := FALSE; udiLastID := 0; uiTargetBand := 0;
	stStatus.udiAcceptedID := 0; stStatus.udiCompletedID := 0;
	tonNoSensor(IN := FALSE);
	tonTravel(IN := FALSE);
END_IF

(* ===== 2. 传感器取反与逐缸姿态判定 ===== *)
aRetract[1] := xSensorRetract1 XOR xInvertSensors;
aExtend[1] := xSensorExtend1 XOR xInvertSensors;
aRetract[2] := xSensorRetract2 XOR xInvertSensors;
aExtend[2] := xSensorExtend2 XOR xInvertSensors;
aRetract[3] := xSensorRetract3 XOR xInvertSensors;
aExtend[3] := xSensorExtend3 XOR xInvertSensors;

(* 单缸两端同时有信号：传感器短路、磁环位置错或机械卡在中间，该缸姿态不可信，按 3003 暴露。
   逐缸判定而不是整组判定：只要有一个缸自相矛盾，整组位置就不可信。 *)
FOR i := 1 TO 3 DO
	IF aRetract[i] AND aExtend[i] THEN
		stStatus.xError := TRUE; stStatus.udiErrorID := 3003;
	END_IF
END_FOR

(* 三缸姿态是否都已确立：每个缸必须恰好一端有效，中间态或两端全无都算未确立。 *)
xAllRetract := aRetract[1] AND aRetract[2] AND aRetract[3];
xPositionKnown := TRUE;
FOR i := 1 TO 3 DO
	IF (NOT aRetract[i]) AND (NOT aExtend[i]) THEN xPositionKnown := FALSE; END_IF
END_FOR
IF stStatus.xError THEN xPositionKnown := FALSE; END_IF

(* 六个传感器全部无信号并持续 tSensorTimeout：判整组传感器丢失，报 3004。
   单缸丢失不在这里报，由 xPositionKnown 为 FALSE 阻断就绪，交给超时暴露，避免一缸调试刷整组报警。 *)
tonNoSensor(IN := xUseReal AND NOT aRetract[1] AND NOT aExtend[1]
	AND NOT aRetract[2] AND NOT aExtend[2]
	AND NOT aRetract[3] AND NOT aExtend[3], PT := tSensorTimeout);
IF tonNoSensor.Q AND NOT stStatus.xError THEN
	stStatus.xError := TRUE; stStatus.udiErrorID := 3004;
END_IF

(* ===== 3. 命令接收与保位判定 ===== *)
IF NOT xUseReal THEN
	(* 未接管：不驱动阀，也不发布就绪，避免被上层当成可用设备 *)
	xCmdValid := FALSE; xTravelling := FALSE; udiLastID := 0; uiTargetBand := 0;
	stStatus.xReady := FALSE; stStatus.xBusy := FALSE; stStatus.xActive := FALSE;
	stStatus.udiAcceptedID := 0; stStatus.udiCompletedID := 0;
ELSIF NOT xEnable OR stStatus.xError OR xFaultHold THEN
	(* 故障或整机故障保持时阀失电，不带错误继续动作 *)
	xCmdValid := FALSE; xTravelling := FALSE;
	stStatus.xReady := FALSE; stStatus.xBusy := FALSE; stStatus.xActive := FALSE;
ELSE
	stStatus.xReady := xEnable AND xPositionKnown;

	(* 新序号即新命令；姿态未确立时不接受，防止朝未知状态动作 *)
	IF (stCommand.udiID <> 0) AND (stCommand.udiID <> udiLastID)
		AND xEnable AND xPositionKnown AND NOT stStatus.xBusy THEN
		udiLastID := stCommand.udiID;
		stStatus.udiAcceptedID := udiLastID; stStatus.udiCompletedID := 0;
		CASE stCommand.eAction OF
		E_DeviceAction.Position:
			IF (stCommand.lrTarget > 0.5) AND (stCommand.lrTarget <= 1.0) THEN
				(* 单缸旧语义：1 = 降到当前料型；料型非法时报 2001，不猜一个缸去动作 *)
				IF (uiMaterialModel = 300) OR (uiMaterialModel = 450) OR (uiMaterialModel = 600) THEN
					uiTargetBand := uiMaterialModel;
				ELSE
					stStatus.xError := TRUE; stStatus.udiErrorID := 2001;
				END_IF
			ELSIF ABS(stCommand.lrTarget) < 0.01 THEN
				uiTargetBand := 0;
			ELSIF (ABS(stCommand.lrTarget - 300.0) < 0.01) THEN
				uiTargetBand := 300;
			ELSIF (ABS(stCommand.lrTarget - 450.0) < 0.01) THEN
				uiTargetBand := 450;
			ELSIF (ABS(stCommand.lrTarget - 600.0) < 0.01) THEN
				uiTargetBand := 600;
			ELSE
				(* 只支持 0 / 300 / 450 / 600，其它目标明确报错而不是静默不动 *)
				stStatus.xError := TRUE; stStatus.udiErrorID := 2001;
			END_IF
			IF NOT stStatus.xError THEN
				xCmdValid := TRUE;
				xTravelling := TRUE;
				stStatus.xBusy := TRUE;
			ELSE
				xCmdValid := FALSE;
			END_IF
		E_DeviceAction.Stop, E_DeviceAction.None:
			xCmdValid := FALSE; xTravelling := FALSE; uiTargetBand := 0;
			stStatus.udiAcceptedID := 0; stStatus.udiCompletedID := 0;
			udiLastID := 0;
		ELSE
			(* 气缸组没有连续运行、点动和回零，明确报错而不是静默不动 *)
			stStatus.xError := TRUE; stStatus.udiErrorID := 2001;
			xCmdValid := FALSE;
		END_CASE
	END_IF

	(* 命令被撤销或失能：立即取消保位，阀随之失电 *)
	IF (stCommand.eAction = E_DeviceAction.Stop) OR (stCommand.eAction = E_DeviceAction.None)
		OR NOT xEnable THEN
		xCmdValid := FALSE; xTravelling := FALSE;
		stStatus.xBusy := FALSE;
	END_IF

	(* 到位判定：目标缸下降到位，并且另外两个缸都在提升位，才算本次命令完成。
	   中间态（目标缸还没下去、或另一缸还没起来）都视为未完成，由超时兜底。 *)
	IF xCmdValid AND xPositionKnown THEN
		CASE uiTargetBand OF
		0:
			IF xAllRetract THEN
				IF xTravelling THEN stStatus.udiCompletedID := udiLastID; END_IF
				xTravelling := FALSE;
				stStatus.xBusy := FALSE;
			END_IF
		300:
			IF aExtend[1] AND aRetract[2] AND aRetract[3] THEN
				IF xTravelling THEN stStatus.udiCompletedID := udiLastID; END_IF
				xTravelling := FALSE;
				stStatus.xBusy := FALSE;
			END_IF
		450:
			IF aExtend[2] AND aRetract[1] AND aRetract[3] THEN
				IF xTravelling THEN stStatus.udiCompletedID := udiLastID; END_IF
				xTravelling := FALSE;
				stStatus.xBusy := FALSE;
			END_IF
		600:
			IF aExtend[3] AND aRetract[1] AND aRetract[2] THEN
				IF xTravelling THEN stStatus.udiCompletedID := udiLastID; END_IF
				xTravelling := FALSE;
				stStatus.xBusy := FALSE;
			END_IF
		END_CASE
	END_IF
END_IF

(* ===== 4. 位置反馈：只有确切在位才更新，中间态保持上次值 ===== *)
IF uiTargetBand = 0 THEN
	IF xAllRetract THEN stStatus.lrPosition := 0.0; END_IF
ELSIF uiTargetBand = 300 THEN
	IF aExtend[1] THEN stStatus.lrPosition := 1.0; END_IF
ELSIF uiTargetBand = 450 THEN
	IF aExtend[2] THEN stStatus.lrPosition := 1.0; END_IF
ELSIF uiTargetBand = 600 THEN
	IF aExtend[3] THEN stStatus.lrPosition := 1.0; END_IF
END_IF

(* 实际下降的料型：命令目标有效且该缸确实到位才报带号，避免阀已得电但没下去时谎报挡料就位 *)
uiActiveBand := 0;
IF (uiTargetBand = 300) AND aExtend[1] THEN uiActiveBand := 300; END_IF
IF (uiTargetBand = 450) AND aExtend[2] THEN uiActiveBand := 450; END_IF
IF (uiTargetBand = 600) AND aExtend[3] THEN uiActiveBand := 600; END_IF

(* ===== 5. 到位超时 ===== *)
tonTravel(IN := xUseReal AND xTravelling AND xCmdValid, PT := tTravelTimeout);
IF tonTravel.Q AND NOT stStatus.xError THEN
	stStatus.xError := TRUE; stStatus.udiErrorID := 3005;
	stStatus.xBusy := FALSE;
	xTravelling := FALSE;
END_IF

(* ===== 6. 阀输出：按保位命令持续输出，不是只在动作过程中输出；任何时刻最多一个缸下降 ===== *)
aValve[1] := FALSE; aValve[2] := FALSE; aValve[3] := FALSE;
IF xCmdValid AND xUseReal AND NOT stStatus.xError AND NOT xFaultHold THEN
	aValve[1] := (uiTargetBand = 300);
	aValve[2] := (uiTargetBand = 450);
	aValve[3] := (uiTargetBand = 600);
END_IF
IF xInvertValve THEN
	aValve[1] := NOT aValve[1]; aValve[2] := NOT aValve[2]; aValve[3] := NOT aValve[3];
END_IF

(* ===== 7. 收尾 ===== *)
stStatus.xReady := stStatus.xReady AND xUseReal AND NOT stStatus.xError;
stStatus.xActive := xCmdValid;
(* 气缸组没有回零动作，用「三缸姿态都已确立」代替，供整机统计已接管设备是否可信 *)
stStatus.xHomed := xUseReal AND xPositionKnown;

(* ---- FB_RealSensor.st ---- *)
FUNCTION_BLOCK FB_RealSensor
(* 模块说明：真实传感器（光电/接近开关）只读适配层。本块不驱动任何输出，只把原始电平
   去抖后发布成「到位」状态，使上层（自动送料判断、互锁、诊断）与仿真设备使用同一套接口。
   按料型/来料判断的是「有没有件」而不是「走到哪个位置」，所以姿态只有 0.0 / 1.0 两端：
   1.0 = 有料（光电被遮挡），0.0 = 无料。连续位置对传感器没有意义。 *)
VAR_INPUT
	xUseReal : BOOL; (* TRUE 表示本编号由真实传感器接管；FALSE 时不读物理点，也不发布就绪。 *)
	xEnable : BOOL; (* 设备级使能，来自整机许可；FALSE 时状态复位为无料且不发布就绪。 *)
	xReset : BOOL; (* 故障复位上升沿；清锁存错误。 *)
	xSensorRaw : BOOL; (* 传感器原始电平，TRUE 表示被遮挡（有料）。 *)
	xInvertSensor : BOOL; (* TRUE 表示接线为低电平有效（遮挡时读 FALSE），本层统一取反，不动上层。 *)
	tDebounce : TIME := T#20MS; (* 去抖时间：光电受粉尘、振动、反光影响会抖，短于该时间的跳变忽略。 *)
	tStuckTimeout : TIME := T#0MS; (* 常亮/常灭监视；0 表示不监视。料走完仍长时间有信号通常代表传感器卡死或反光。 *)
	stConfig : ST_DeviceConfig; (* 与其它设备一致的配置结构；传感器只用 lrInitialPosition 作初值，不使用行程字段。 *)
	stCommand : ST_DeviceCommand; (* 上层统一设备命令；传感器只响应被读请求，Position 目标被忽略。 *)
END_VAR
VAR_OUTPUT
	stStatus : ST_DeviceStatus; (* 与仿真侧语义一致；lrPosition 取 1.0 有料、0.0 无料。 *)
	xDetected : BOOL; (* 去抖后的最终信号，TRUE=有料。流程与互锁直接取用这个而不是原始点。 *)
	xRaw : BOOL; (* 取反处理后的原始电平（未去抖），供在线排查接线极性与抖动。 *)
END_VAR
VAR
	rtReset : R_TRIG; (* 复位上升沿。 *)
	tonDebounce : TON; (* 由 FALSE 变 TRUE 的去抖计时，到时才认「有料」。 *)
	tonClear : TON; (* 由 TRUE 变 FALSE 的去抖计时，到时才认「无料」。 *)
	tonStuck : TON; (* 长时间保持同一状态计时，用于常亮/常灭监视。 *)
	xStuckWindowClear : BOOL; (* 本扫描检测到电平跳变：清掉常亮/常灭计时窗口，重新开始计时。 *)
	xStable : BOOL; (* 去抖后的稳定值。 *)
	xLastRaw : BOOL; (* 上扫描取反后的原始电平，用于判断是否发生跳变并重置去抖计时。 *)
	xBooted : BOOL; (* 首次扫描标志，上电时直接用当前电平作初值，不等待去抖。 *)
END_VAR
FUNCTION_BLOCK FB_RealSensor
rtReset(CLK := xReset);

(* ===== 1. 复位：只清错误，状态仍由传感器决定 ===== *)
IF xUseReal AND rtReset.Q THEN
	stStatus.xError := FALSE; stStatus.udiErrorID := 0;
	tonStuck(IN := FALSE);
END_IF

(* ===== 2. 极性处理：接线反了只改 xInvertSensor 一个参数，上层不受影响 ===== *)
xRaw := xSensorRaw XOR xInvertSensor;

(* ===== 3. 去抖：跳变后必须稳定 tDebounce 才改 xStable ===== *)
(* 用两个单稳计时而不是一个沿检测，是为了让"抖动期间保持上次稳定值"这件事显式可见：
   信号连续抖动时两个计时都不会到时，xStable 保持在最后一个稳定值上。 *)
xStuckWindowClear := (NOT xBooted) OR (xRaw <> xLastRaw);
IF xStuckWindowClear THEN
	tonDebounce(IN := FALSE);
	tonClear(IN := FALSE);
	IF NOT xBooted THEN
		(* 上电直接用当前电平作初值，避免开机 20ms 内把有料当无料 *)
		xStable := xRaw;
		xBooted := TRUE;
	END_IF
	xLastRaw := xRaw;
END_IF

IF xUseReal THEN
	IF xRaw THEN
		tonDebounce(IN := TRUE, PT := tDebounce);
		tonClear(IN := FALSE);
		IF tonDebounce.Q THEN xStable := TRUE; END_IF
	ELSE
		tonClear(IN := TRUE, PT := tDebounce);
		tonDebounce(IN := FALSE);
		IF tonClear.Q THEN xStable := FALSE; END_IF
	END_IF
END_IF

xDetected := xStable;

(* ===== 4. 常亮/常灭监视：料已走完却一直有信号，或本该有料却一直没有，都报出来 =====
   只监视"信号纹丝不动"这个可观测事实，不猜业务含义；阈值由 tStuckTimeout 给，0 表示关闭。 *)
tonStuck(IN := xUseReal AND (tStuckTimeout > T#0MS) AND NOT xStuckWindowClear, PT := tStuckTimeout);
IF tonStuck.Q AND NOT stStatus.xError THEN
	stStatus.xError := TRUE;
	(* 3006：持续有信号（常亮/反光/卡死）；3007：持续无信号（断线/被挡/未接通） *)
	IF xDetected THEN stStatus.udiErrorID := 3006;
	ELSE stStatus.udiErrorID := 3007; END_IF
END_IF

(* ===== 5. 状态发布：传感器没有动作请求，只要接管且使能就算就绪 ===== *)
stStatus.lrPosition := SEL(xDetected, 0.0, 1.0);
stStatus.xReady := xUseReal AND xEnable AND NOT stStatus.xError;
stStatus.xActive := xUseReal AND xDetected;
stStatus.xBusy := FALSE;
(* 传感器没有回零概念，用"已接管且状态可信"代替 *)
stStatus.xHomed := xUseReal AND xBooted;
stStatus.xRealActive := xUseReal;

(* ---- FB_Valve.st ---- *)
(* 模块说明：阀适配入口，供喷油 G5 和吹气 G6 使用。当前用运行状态表示开启，未映射输出。 *)
FUNCTION_BLOCK FB_Valve
VAR_INPUT
    xSimulation : BOOL; (* TRUE 使用内部仿真；当前 FALSE 报未实现 3001，不会接管真实运动。 *)
    xEnable : BOOL; (* 本功能使能，电平有效；失能时不接受新的动作请求。 *)
    xReset : BOOL; (* 故障复位许可；仿真设备仅在故障注入已撤销时清除错误。 *)
    xStall : BOOL; (* 仿真卡住输入；TRUE 暂停位置推进且不发完成，保留忙状态。 *)
    xInjectFault : BOOL; (* 仿真设备故障输入；TRUE 锁存错误码 9001。 *)
    stConfig : ST_DeviceConfig; (* 设备类型、初始位置、软限位与仿真动作时间。 *)
    stCommand : ST_DeviceCommand; (* 当前单设备命令，含动作类型、序号、目标和速度。 *)
END_VAR
VAR_OUTPUT
    stStatus : ST_DeviceStatus; (* 本模块对外发布的状态；字段含义见其数据类型。 *)
END_VAR
VAR
    fbSimulation : FB_SimDevice; (* 内部设备仿真实例，真实设备适配尚未接入。 *)
END_VAR
FUNCTION_BLOCK FB_Valve
(* 真实设备适配尚未接入；关闭仿真时返回 3001，避免误认为已具备实机控制。 *)
fbSimulation(xEnable := xEnable AND xSimulation, xReset := xReset,
    xStall := xStall, xInjectFault := xInjectFault,
    stConfig := stConfig, stCommand := stCommand);
stStatus := fbSimulation.stStatus;
IF NOT xSimulation THEN
    stStatus.xReady := FALSE; stStatus.xBusy := FALSE; stStatus.xActive := FALSE;
    stStatus.xError := TRUE; stStatus.udiErrorID := 3001;
END_IF
